Fanuc KAREL source: KT00419.KL

PROGRAM KT00419
%NOLOCKGROUP
VAR
  P1: POSITION
  P2: POSITION
  OUT: BOOLEAN
BEGIN
  OUT = P1 > P2
END KT00419
